(* IEC 61131-3 sources: llm-plc-st-eval/data/processed/gpt-4o/B3/zero_shot, 3 files *)

(* ---- ejec_1.st ---- *)
FUNCTION_BLOCK FB_Contador
VAR_INPUT
    sensorPieza : BOOL;  // Entrada del sensor fotoeléctrico
    btnReset : BOOL;     // Botón de reset
END_VAR

VAR_OUTPUT
    loteListo : BOOL;    // Indica si el lote está completo
    cuenta : INT;        // Contador de piezas
END_VAR

VAR
    prevSensorPieza : BOOL;  // Estado anterior del sensor
END_VAR

// Inicialización de variables
IF btnReset THEN
    cuenta := 0;         // Reinicia el contador
    loteListo := FALSE;  // Desactiva la salida de lote completo
ELSE
    // Detecta el flanco ascendente del sensor
    IF (sensorPieza AND NOT prevSensorPieza) THEN
        cuenta := cuenta + 1;  // Incrementa el contador
    END_IF

    // Verifica si el lote está completo
    IF cuenta >= 12 THEN
        loteListo := TRUE;  // Activa la salida de lote completo
    ELSE
        loteListo := FALSE; // Asegura que la salida esté desactivada si no está completo
    END_IF
END_IF

// Actualiza el estado anterior del sensor
prevSensorPieza := sensorPieza;

END_FUNCTION_BLOCK

(* ---- ejec_2.st ---- *)
FUNCTION_BLOCK FB_Contador
VAR_INPUT
    sensorPieza : BOOL;  // Sensor que detecta la pieza
    btnReset : BOOL;     // Botón para resetear el contador
END_VAR

VAR_OUTPUT
    loteListo : BOOL;    // Indica si el lote está completo
    cuenta : INT;        // Contador de piezas
END_VAR

VAR
    prevSensorPieza : BOOL;  // Estado previo del sensor
END_VAR

// Inicialización de variables
INIT
    cuenta := 0;
    loteListo := FALSE;
    prevSensorPieza := FALSE;
END_INIT

// Cuerpo del bloque de función
IF btnReset THEN
    // Si el botón de reset está presionado, reiniciar el contador y la salida de lote
    cuenta := 0;
    loteListo := FALSE;
ELSIF NOT prevSensorPieza AND sensorPieza THEN
    // Detectar flanco ascendente del sensor
    cuenta := cuenta + 1;
    IF cuenta >= 12 THEN
        // Si se han contado 12 piezas, activar la salida de lote completo
        loteListo := TRUE;
    END_IF
END_IF

// Actualizar el estado previo del sensor
prevSensorPieza := sensorPieza;

END_FUNCTION_BLOCK

(* ---- ejec_3.st ---- *)
FUNCTION_BLOCK FB_Contador
VAR_INPUT
    sensorPieza : BOOL;  // Entrada del sensor fotoeléctrico
    btnReset : BOOL;     // Botón de reset
END_VAR

VAR_OUTPUT
    loteListo : BOOL;    // Salida que indica si el lote está completo
    cuenta : INT;        // Contador de piezas
END_VAR

VAR
    prevSensorPieza : BOOL;  // Estado anterior del sensor
END_VAR

// Inicialización de variables
IF btnReset THEN
    cuenta := 0;         // Reinicia el contador
    loteListo := FALSE;  // Desactiva la salida de lote completo
END_IF

// Detección de flanco ascendente del sensor
IF (sensorPieza AND NOT prevSensorPieza) THEN
    cuenta := cuenta + 1;  // Incrementa el contador
END_IF

// Verificación de lote completo
IF cuenta >= 12 THEN
    loteListo := TRUE;  // Activa la salida de lote completo
ELSE
    loteListo := FALSE; // Asegura que la salida esté desactivada si no se completa el lote
END_IF

// Actualización del estado anterior del sensor
prevSensorPieza := sensorPieza;

END_FUNCTION_BLOCK
